Fanuc KAREL source: kt00081.KL

-- PROVISIONAL review KL for V940-1; original PC SHA256 174a0ffbc7c028999a94cc4052265e6b4a995addd64d243aa7130bd31d446019
-- Incomplete behavior may be omitted. Consult companion uncertainty JSON. Do not deploy.
PROGRAM KT00081
%NOLOCKGROUP
VAR
  I2 : INTEGER
  OUT : INTEGER
-- UNRESOLVED_DECL Y1 type=002018
BEGIN
  -- V9_ZERO_TABLE_METADATA_HINT layout=0001; no indexed target words; source/name/runtime held
  -- UNRESOLVED_PC offsets 5-19; opcodes 2E,22,9D,33,B2
  -- UNRESOLVED_PC offsets 24-35; opcodes 2E,23
  -- UNRESOLVED_PC offsets 40-62; opcodes 22,9D,33,B1,21,54,23
  -- UNRESOLVED_PC offsets 67-71; opcodes 7F
END KT00081
